(* IEC 61131-3 sources: Test-Git_ESME26/TestProgettoESME_26.fbsproj/PacDriveLib Migration/Motion/PDL_FB_PosOnTorque.fb.st^, 2 files *)

(* ---- InitInterfaces.meth.st ---- *)
METHOD InitInterfaces : BOOL
VAR_INPUT
END_VAR

	IF i_ifDrive = 0 THEN
		q_etDiag	:= GD.ET_Diag.InputParameterInvalid;
		q_etDiagExt := PDL_ET_DiagExt.DriveInvalid;
		q_sMsg		:= 'i_ifDrive - Invalid Interface';
		RETURN;
	END_IF

	xSuccess := __QUERYINTERFACE(i_ifDrive, ifGetParentDevice);
	IF NOT xSuccess OR ifGetParentDevice = 0 THEN
		q_etDiag	:= GD.ET_Diag.InputParameterInvalid;
		q_etDiagExt := PDL_ET_DiagExt.DriveInvalid;
		q_sMsg		:= 'i_ifDrive - IF_GetParentDevice not implemented.';
		RETURN;
	END_IF
	ifDeviceAccess := ifGetParentDevice.GetParentDevice();

	xSuccess := __QUERYINTERFACE(ifDeviceAccess,ifDriveConfigAccess );
	IF (NOT xSuccess OR ifDriveConfigAccess = 0) THEN
		q_etDiag	:= GD.ET_Diag.InputParameterInvalid;
		q_etDiagExt := PDL_ET_DiagExt.DriveInvalid;
		q_sMsg		:= 'i_ifDrive - IF_DriveConfig not implemented.';
		diState := 0;
		RETURN;
	END_IF
	ifDriveConfig := ifDriveConfigAccess.DriveConfig;

	xSuccess := __QUERYINTERFACE(ifDeviceAccess,ifDriveCurrentAccess );
	IF (NOT xSuccess OR ifDriveCurrentAccess = 0) THEN
		q_etDiag	:= GD.ET_Diag.InputParameterInvalid;
		q_etDiagExt := PDL_ET_DiagExt.DriveInvalid;
		q_sMsg		:= 'i_ifDrive - IF_DriveCurrent not implemented.';
		diState := 0;
		RETURN;
	END_IF
	ifDriveCurrent := ifDriveCurrentAccess.DriveCurrent;

	xSuccess := __QUERYINTERFACE(ifDeviceAccess,ifDriveAccess );
	IF (NOT xSuccess OR ifDriveAccess = 0) THEN
		q_etDiag	:= GD.ET_Diag.InputParameterInvalid;
		q_etDiagExt := PDL_ET_DiagExt.DriveInvalid;
		q_sMsg		:= 'i_ifDrive - IF_Drive not implemented.';
		diState := 0;
		RETURN;
	END_IF
	ifDrive := ifDriveAccess.Drive;

	xSuccess := __QUERYINTERFACE(ifDeviceAccess,ifMotorAccess );
	IF (NOT xSuccess OR ifMotorAccess = 0) THEN
		q_etDiag	:= GD.ET_Diag.InputParameterInvalid;
		q_etDiagExt := PDL_ET_DiagExt.DriveInvalid;
		q_sMsg		:= 'i_ifDrive - IF_Motor not implemented.';
		diState := 0;
		RETURN;
	END_IF
	ifMotor := ifMotorAccess.Motor;

(* ---- lrMaxPossibleTorque.prop.st ---- *)
PROPERTY lrMaxPossibleTorque : LREAL
__GETTERDECLARATION__
VAR
END_VAR
__GETTERIMPLEMENTATION__
lrMaxPossibleTorque := lrMaxPossibleTorque_loc;
